// TwinCAT 3 PLC project ArbiterPLC
// ProgramVersion: 3.1.4022.7
// libraries:
//   LCLS General, * (SLAC)
//   Tc2_MC2, * (Beckhoff Automation GmbH)
//   Tc2_Standard, * (Beckhoff Automation GmbH)
//   Tc2_System, * (Beckhoff Automation GmbH)
//   Tc2_SystemCX, * (Beckhoff Automation GmbH)
//   Tc2_Utilities, * (Beckhoff Automation GmbH)
//   Tc3_Module, * (Beckhoff Automation GmbH)
//   PMPS,0.0.0,SLAC - LCLS
// project tree:
//   / FFOTask.TcTTO, PlcTask.TcTTO
//   GVLs/ GVL.TcGVL, GVL_CheckBounds.TcGVL
//   ImplicitChecks/ CheckBounds.TcPOU, CheckRangeSigned.TcPOU, CheckRangeUnsigned.TcPOU
//   POUs/ Fast_Faults_Evaluate.TcPOU, FB_eVSimulator.TcPOU, FB_SubSystem_PMPS_IO.TcPOU, MachineSimulation.TcPOU, MAIN.TcPOU, PMPS_Arbiter.TcPOU
// real-time tasks:
//   TASK PlcTask: cycle T#10ms, priority 2, ADS port 350
//   TASK FFOTask: cycle T#1ms, priority 1, ADS port 351
// I/O:
//   DEVICE Device 1 (EtherCAT), AmsNetId 0.0.0.0.2.1
//     Term 1 (EK1200) [EK1200-5000 EtherCAT Power supply (2A E-Bus)]
//       PMPS_FFO [EL2022 2Ch. Dig. Output 24V, 2A]
//       PMPS_BC [EL2809 16Ch. Dig. Output 24V, 0.5A]
//       PMPS_CLTS [EL2809 16Ch. Dig. Output 24V, 0.5A]
//       Term 3 (EK1122) [EK1122 2 port EtherCAT junction]
//         SubSysPLC1 [EL6692 EtherCAT Bridge terminal (Secondary)]
//         SubSysPLC2 [EL6692 EtherCAT Bridge terminal (Secondary)]
//       Term 6 (EK1110) [EK1110 EtherCAT extension]
// variable links:
//   ArbiterPLC Instance <-> Device 1 (EtherCAT)/Term 1 (EK1200)/PMPS_BC
//     PlcTask Outputs/PMPS_Arbiter.fbMPSInterface.q_BC_ASSERTION_LINES[{1..16}] <-> Channel {1..16}/Output  (16 links)
//   ArbiterPLC Instance <-> Device 1 (EtherCAT)/Term 1 (EK1200)/PMPS_CLTS
//     PlcTask Outputs/PMPS_Arbiter.fbCuInterface.q_CLTS_ASSERTION_LINES[{1..16}] <-> Channel {1..16}/Output  (16 links)
//   ArbiterPLC Instance <-> Device 1 (EtherCAT)/Term 1 (EK1200)/PMPS_FFO
//     FFOTask Outputs/GVL.g_FastFaultOutput1.q_xFastFaultOut <-> Channel 1/Output
//   ArbiterPLC Instance <-> Device 1 (EtherCAT)/Term 1 (EK1200)/Term 3 (EK1122)/SubSysPLC1
//     PlcTask Inputs/PMPS_Arbiter.fbSubSys1_PMPS_IO.i_Connected <-> SYNC Inputs/External device not connected
//     PlcTask Inputs/PMPS_Arbiter.fbSubSys1_PMPS_IO.i_RequestedBP <-> IO Inputs/RequestedBP
//     PlcTask Inputs/PMPS_Arbiter.fbSubSys1_PMPS_IO.i_TxPDOState <-> SYNC Inputs/TxPDO state
//     PlcTask Inputs/PMPS_Arbiter.fbSubSys1_PMPS_IO.i_WcState <-> WcState/WcState
//     PlcTask Outputs/PMPS_Arbiter.fbSubSys1_PMPS_IO.o_CurrentBP <-> IO Outputs/CurrentBP
//   ArbiterPLC Instance <-> Device 1 (EtherCAT)/Term 1 (EK1200)/Term 3 (EK1122)/SubSysPLC2
//     PlcTask Inputs/PMPS_Arbiter.fbSubSys2_PMPS_IO.i_Connected <-> SYNC Inputs/External device not connected
//     PlcTask Inputs/PMPS_Arbiter.fbSubSys2_PMPS_IO.i_RequestedBP <-> IO Inputs/RequestedBP
//     PlcTask Inputs/PMPS_Arbiter.fbSubSys2_PMPS_IO.i_TxPDOState <-> SYNC Inputs/TxPDO state
//     PlcTask Inputs/PMPS_Arbiter.fbSubSys2_PMPS_IO.i_WcState <-> WcState/WcState
//     PlcTask Outputs/PMPS_Arbiter.fbSubSys2_PMPS_IO.o_CurrentBP <-> IO Outputs/CurrentBP

CONFIGURATION ArbiterPLC
    RESOURCE PLC ON TwinCAT3
        TASK FFOTask(INTERVAL := T#1ms, PRIORITY := 1);
        TASK PlcTask(INTERVAL := T#10ms, PRIORITY := 2);
        PROGRAM Fast_Faults_Evaluate WITH FFOTask : Fast_Faults_Evaluate;
        PROGRAM MAIN WITH PlcTask : MAIN;
    END_RESOURCE
END_CONFIGURATION

// ---- GVLs/GVL.TcGVL

VAR_GLOBAL
   {attribute 'pytmc' := '
    pv: ARBITER:K:Arbiter1
    '}
	g_fbArbiter1	:	FB_Arbiter;

	ReqBP	:	ST_BeamParams; //Currently the placeholder for the fully arbitrated BP set
	
	//Example implementation of the FFO
    (*
    {attribute 'pytmc' := '
    pv: ARBITER:K:FF1
    '} *)
	{attribute 'TcLinkTo' := '.q_xFastFaultOut:=TIIB[PMPS_FFO]^Channel 1^Output'}
	g_FastFaultOutput1	:	FB_HardwareFFOutput;
    
	g_rTestingVelocity	:	LREAL := PMPS_GVL.VISIBLE_TEST_VELOCITY;
    
    AttemptReset    :   BOOL; // For testing
END_VAR

// ---- GVLs/GVL_CheckBounds.TcGVL
{attribute 'qualified_only'}
VAR_GLOBAL
    nTooLow : UDINT;
    nTooHigh : UDINT;
    nDivByZero : UDINT;
END_VAR

// ---- POUs/Fast_Faults_Evaluate.TcPOU
PROGRAM Fast_Faults_Evaluate
VAR
END_VAR

g_FastFaultOutput1.EvaluateOutput();

END_PROGRAM

// ---- POUs/MAIN.TcPOU
PROGRAM MAIN
VAR
	Initialize	:	BOOL := TRUE;
	
	AttemptReset : TON := (PT:=T#500ms);
    
    DisplayStats : FB_CXSetTextDisplayUSB := (nPort:=28928);
    fbFormat   : FB_FormatString;
    bError     : BOOL;
    nErrID     : UDINT;
    sOut       : T_MaxString;   

END_VAR

//Arbiter PLC

IF Initialize THEN

	g_fbArbiter1.A_Init();

	Initialize := FALSE;
END_IF

MachineSimulation();
		
PMPS_Arbiter();


AttemptReset(IN:=GVL.g_FastFaultOutput1.xOK, Q=>GVL.g_FastFaultOutput1.i_xReset);


DisplayStats.bExecute S= NOT DisplayStats.bBusy AND NOT DisplayStats.bError;
DisplayStats.bExecute R= DisplayStats.bBusy OR DisplayStats.bError;

DisplayStats.sLine1 := 'PMPS-ARBITER-K';
fbFormat(sFormat := 'Fast Faults: %d', arg1:=F_ULINT(PMPS_GVL.AccumulatedFF), sOut=>DisplayStats.sLine2, bError => bError, nErrID => nErrID ); 

DisplayStats(eMode:=E_CX2100_DisplayModesWr.eCX2100_WriteLines);

ACTION Initialize:

END_ACTION

END_PROGRAM

// ---- POUs/MachineSimulation.TcPOU
PROGRAM MachineSimulation
VAR
	fbMachine	:	FB_MachineSimulator; //Simulates attenuator as well
	fbeVSimulator : FB_eVSimulator := (NoiseLevel := 1);
END_VAR

// reV Simulator
fbeVSimulator(eV => fbMachine.i_reV);

// Machine simulator
fbMachine(
	i_stAssertedParams := ReqBP,
	q_stMachineParams => PMPS_GVL.stCurrentBeamParameters,
	i_xFault	:= NOT GVL.g_FastFaultOutput1.q_xFastFaultOut
	);

PMPS_GVL.stCurrentBeamParameters.neVRange := F_eVRangeCalculator(fbMachine.q_stMachineParams.reV, PMPS_GVL.stCurrentBeamParameters.neVRange);

END_PROGRAM

// ---- POUs/FB_eVSimulator.TcPOU
(* eV Simulator
A. Wallace 2019-8-30

Adds noise to the eV and changes eV position occasionally.
*)
FUNCTION_BLOCK FB_eVSimulator
VAR_INPUT
	NoiseLevel	:	REAL	:= 0; // eV Noise
	ChangeTime : TIME := T#10S;
END_VAR
VAR_OUTPUT
	eV	:	REAL := 300;
END_VAR
VAR
	eVRange : REAL := 1600;
	timer: TON;
	eVRand	:	DRAND :=(Seed:=0);
	NoiseRand : DRAND := (Seed:=0);
END_VAR


timer(in:=TRUE, PT:=ChangeTime);

//Occasionally change eV
IF timer.Q THEN
	timer(in:=FALSE);
	eVRand();
	eV := LIMIT(0, eVRange*LREAL_TO_REAL(eVRand.Num), eVRange);
END_IF

// Noise generation
NoiseRand();
eV := eV + NoiseLevel*LREAL_TO_REAL(NoiseRand.Num);
NoiseRand();
eV := LIMIT(0, ev - NoiseLevel*LREAL_TO_REAL(NoiseRand.Num), eVRange);

END_FUNCTION_BLOCK

// ---- POUs/PMPS_Arbiter.TcPOU
PROGRAM PMPS_Arbiter
VAR
	
	fbPhotonEnergyWatcher	:	FB_PhotonEnergyWatcher;
	
	fbMPSInterface	:	FB_BeamClassOutputs;
    
    fbCuInterface	:	FB_CTLS_Outputs;
	
	(* Subsystem requests use this FB and a pragma link to pass their requests to the arbiter.
	The fb is called on each cycle and updates the arbiter with the current BP set requested 
	from the subsystem PLC.*)
	//<TODO> make this so it does input and output to the IF
	{attribute 'TcLinkTo' := '.i_RequestedBP:=TIIB[SubSysPLC1]^IO Inputs^RequestedBP; 
                                .o_CurrentBP:=TIIB[SubSysPLC1]^IO Outputs^CurrentBP;
                                .i_Connected:=TIIB[SubSysPLC1]^SYNC Inputs^External device not connected;
                                .i_WcState:=TIIB[SubSysPLC1]^WcState^WcState;
                                .i_TxPDOState:=TIIB[SubSysPLC1]^SYNC Inputs^TxPDO state;
                                '}
	fbSubSys1_PMPS_IO : FB_SubSystem_PMPS_IO := (RequestingSystemID := 16#FF0F);
	
	{attribute 'TcLinkTo' := '.i_RequestedBP:=TIIB[SubSysPLC2]^IO Inputs^RequestedBP; 
                                .o_CurrentBP:=TIIB[SubSysPLC2]^IO Outputs^CurrentBP;
                                .i_Connected:=TIIB[SubSysPLC2]^SYNC Inputs^External device not connected;
                                .i_WcState:=TIIB[SubSysPLC2]^WcState^WcState;
                                .i_TxPDOState:=TIIB[SubSysPLC2]^SYNC Inputs^TxPDO state;
                                '}
	fbSubSys2_PMPS_IO : FB_SubSystem_PMPS_IO := (RequestingSystemID := 16#FF10);
	
	AttemptReset : TON := (PT:=T#1s);
    
    anothervar : bool;
	
END_VAR


// Updating arbiter with subsystem requests.
fbSubSys1_PMPS_IO(Arbiter:=GVL.g_fbArbiter1, fbFFHWO:=GVL.g_FastFaultOutput1, Reset:=GVL.AttemptReset);

fbSubSys2_PMPS_IO(Arbiter:=GVL.g_fbArbiter1, fbFFHWO:=GVL.g_FastFaultOutput1, Reset:=GVL.AttemptReset);

// Example with attenuator peel-off
//////////////////////////////////

// Beam parameter requestor
ReqBP := g_fbArbiter1.GetArbitratedBP();

// Request beam class
fbMPSInterface(i_ArbiterBP := ReqBP);

// Request Cu beam rate
fbCuInterface(i_ArbiterBP := ReqBP);

// Calculate the current eV word
PMPS_GVL.stCurrentBeamParameters.neVRange := F_eVRangeCalculator(
	PMPS_GVL.stCurrentBeamParameters.reV,
	PMPS_GVL.stCurrentBeamParameters.neVRange);

// Keep an eye on the photon energy
fbPhotonEnergyWatcher(i_stCurrentBeamParams	:= PMPS_GVL.stCurrentBeamParameters,
					i_stRequestedBeamParams := ReqBP,
					io_fbFFHWO:= GVL.g_FastFaultOutput1,
                    i_xReset := GVL.AttemptReset);

AttemptReset(IN:=fbPhotonEnergyWatcher.xPhotonEnergyWithinBounds, Q=>GVL.AttemptReset);

END_PROGRAM

// ---- POUs/FB_SubSystem_PMPS_IO.TcPOU
(* Exchanges preemption requests and current beam state with subsystems in arbiter
network.

2019-12-2, A. Wallace

*)
FUNCTION_BLOCK FB_SubSystem_PMPS_IO
VAR_INPUT
	RequestingSystemID	:	DWORD := PMPS_GVL.EXCLUDED_ASSERTION_ID; // System ID for making requests to the supreme arbiter
    Reset : BOOL;
END_VAR
VAR_OUTPUT
END_VAR
VAR_IN_OUT
	Arbiter	: FB_Arbiter;
    fbFFHWO : FB_HardwareFFOutput;
END_VAR
VAR
	i_RequestedBP AT %I*	:	ST_BeamParams;
	o_CurrentBP AT %Q* : ST_BeamParams;
    
    // EL6692 Diagnostics
    i_Connected AT %I* : BOOL; // SYNC Inputs^External device not connected !!! Doesn't really work.
    i_WcState AT %I* : BOOL; // WcState^WcState
    i_TxPDOState AT %I* : BOOL; // SYNC Inputs^TxPDO state
    
    // Fast faults
    ffPMPSIO_Disconnect : FB_FastFault := (i_Desc:='Fast fault on arbiter disconnection');
END_VAR

// Update arbiter with our request
Arbiter.RemoveRequest(RequestingSystemID);
Arbiter.AddRequest(RequestingSystemID, i_RequestedBP);

// Current beam params fanout
o_CurrentBP := PMPS_GVL.stCurrentBeamParameters;

// Both of these values should be 0 for a fully valid exchange
ffPMPSIO_Disconnect.i_xOK := NOT i_WcState AND NOT i_TxPDOState;

ffPMPSIO_Disconnect(
    io_fbFFHWO := fbFFHWO,
    i_xReset := Reset);

END_FUNCTION_BLOCK

// ---- ImplicitChecks/CheckBounds.TcPOU
// Implicitly generated code : DO NOT EDIT
FUNCTION CheckBounds : DINT
VAR_INPUT
	index, lower, upper: DINT;
END_VAR
// User defined local variables
VAR
    sMessageLow   : STRING := 'CheckBounds: Index too low (%d)';
    sMessageHigh  : STRING := 'CheckBounds: Index too high (%d)';
END_VAR

// Index too low
IF index < lower THEN
    CheckBounds := lower;
    // Increase global counter
    GVL_CheckBounds.nTooLow := GVL_CheckBounds.nTooLow + 1;
    // Log message
    ADSLOGDINT(msgCtrlMask := ADSLOG_MSGTYPE_WARN,
               msgFmtStr   := sMessageLow,
               dintArg     := index);

// Index too high
ELSIF index > upper THEN
    CheckBounds := upper;
    // Increase global counter
    GVL_CheckBounds.nTooHigh := GVL_CheckBounds.nTooHigh + 1;
    // Log message
    ADSLOGDINT(msgCtrlMask := ADSLOG_MSGTYPE_WARN,
               msgFmtStr   := sMessageHigh,
               dintArg     := index);

// Index OK
ELSE 
    CheckBounds := index;
END_IF
{flow}

END_FUNCTION

// ---- ImplicitChecks/CheckRangeSigned.TcPOU
// Implicitly generated code : DO NOT EDIT
FUNCTION CheckRangeSigned : DINT
VAR_INPUT
	value, lower, upper: DINT;
END_VAR

// Implicitly generated code : Only an Implementation suggestion

IF (value < lower) THEN
	CheckRangeSigned := lower;
ELSIF(value > upper) THEN
	CheckRangeSigned := upper;
ELSE
	CheckRangeSigned := value;
END_IF
{flow}

END_FUNCTION

// ---- ImplicitChecks/CheckRangeUnsigned.TcPOU
// Implicitly generated code : DO NOT EDIT
FUNCTION CheckRangeUnsigned : UDINT
VAR_INPUT
	value, lower, upper: UDINT;
END_VAR

// Implicitly generated code : Only an Implementation suggestion
{noflow}
IF (value < lower) THEN
	CheckRangeUnsigned := lower;
ELSIF(value > upper) THEN
	CheckRangeUnsigned := upper;
ELSE
	CheckRangeUnsigned := value;
END_IF
{flow}

END_FUNCTION
